Staubli VAL3: _onStartTRAJ.pgx

public program _onStartTRAJ()
begin
  nPgIndexTRAJ=0
  nPgNumTRAJ=0
  sPageTRAJ=""
  sPgIndexTRAJ=""
//  call resfreshTRAJ()
end
